// TIA Portal project "项目6" (V15.1)

(* hardware
DEVICE "S7-1200 station_1"  S7-1200 Station
   slot 0: "Rack_0"  S7-1200 Rack  Rack  V1.0
   slot 1: "PLC_1"  CPU 1214C DC/DC/DC  6ES7 214-1AG40-0XB0  V4.2
   slot 2: "DI 16/DQ 16x24VDC_1"  6ES7 223-1BL32-0XB0  V2.0
   slot 3: "AI 4x13BIT/AQ 2x14BIT_1"  6ES7 234-4HE32-0XB0  V2.0
DEVICE "HMI_1"  KTP700 Basic PN
   slot 0: "HMI_1"  KTP700 Basic PN  6AV2 123-2GB03-0AX0  15.1.0.0
   slot 1: "HMI_RT_1"  KTP700 Basic PN  6AV2 123-2GB03-0AX0  15.1.0.0
   slot 5: "HMI_1.IE_CP_1"  PROFINET Interface  15.0.1.0
      slot 1: "PROFINET Interface_1"  PROFINET Interface
         slot 1: "Port_1"  Port
*)

// ===== PLC "PLC_1"  CPU 1214C DC/DC/DC =====

VAR_GLOBAL   // PLC tag table "IO变量表"
   "手动自动切换" AT %I9.0 : Bool;
   "点动正转" AT %I9.1 : Bool;
   "点动反转" AT %I9.2 : Bool;
   "自动定位启动" AT %I9.5 : Bool;
   "停止按钮" AT %I9.7 : Bool;
   "电机脉冲" AT %Q0.0 : Bool;
   "电机方向" AT %Q0.1 : Bool;
   "电机使能" AT %Q1.0 : Bool;
   "回原点启动" AT %I0.3 : Bool;
   "循环" AT %I9.6 : Bool;
   "回原点" AT %I9.3 : Bool;
END_VAR

VAR_GLOBAL   // PLC tag table "数据变量表"
   "自动状态" AT %MW10 : Int;
   "B点坐标" AT %MD20 : Real;
   "C点坐标" AT %MD24 : Real;
   "点动速度" AT %MD28 : Real;   // 120-1800
   "自动运行速度" AT %MD32 : Real;   // 120-1800
END_VAR

// folder: System blocks/Program resources

DATA_BLOCK "B点延时_DB"   // DB7
{ S7_Optimized_Access := 'TRUE' }
AUTHOR : Simatic
FAMILY : IEC
NAME : IEC_TMR
VERSION : 1.0
// stored: InstanceOfName IEC_TIMER
"IEC_TIMER"
BEGIN
END_DATA_BLOCK

DATA_BLOCK "C点延时_DB"   // DB8
{ S7_Optimized_Access := 'TRUE' }
AUTHOR : Simatic
FAMILY : IEC
NAME : IEC_TMR
VERSION : 1.0
// stored: InstanceOfName IEC_TIMER
"IEC_TIMER"
BEGIN
END_DATA_BLOCK

// folder: (top level)

DATA_BLOCK "步进电机"   // DB1, Motion_DB
{ S7_Optimized_Access := 'TRUE' }
AUTHOR : SIMATIC
FAMILY : BasicMC
NAME : TO_PosAx
VERSION : 6.0
// stored: InstanceOfName TO_PositioningAxis
"TO_PositioningAxis"
BEGIN
   // Axis.HomingReferencePointSwitch_AddressCU = %I0.3
   // Axis.LengthUnitNormalized.Distance = 1005
   // Axis.EnableOutput_AddressCU = %Q1.0
   // Axis.OnlinePtoModeCU = 16#0000_0002
   // Axis.DirectionOutputEnabledCU = TRUE
   // Axis.SelectedChannel2EnumCU = %Q0.1
   // Axis.SelectedChannel1EnumCU = %Q0.0
   // Pulse.MinDeltaDeltaFrequencyCU = 0.004
   // Pulse.MaxDeltaDeltaFrequencyCU = 1.0E+10
   // Pulse.MinDeltaFrequencyCU = 0.005
   // Pulse.MaxDeltaFrequencyCU = 9.5E+9
   // Pulse.MinFrequencyCU = 1.0
   // Pulse.MaxFrequencyCU = 100000.0
   // Pulse.OutputSourceCU = 16#0000_0000
   // Axis.SelectPTO = 0
   // Axis.LengthUnit.LastDistance = 1005
END_DATA_BLOCK

ORGANIZATION_BLOCK "Main"   // OB1, SCL, ProgramCycle
TITLE = "Main Program Sweep (Cycle)"
{ S7_Optimized_Access := 'TRUE' }
VERSION : 0.1
   VAR_INPUT
      Initial_Call : Bool;   // Initial call of this OB
      Remanence : Bool;   // =True, if remanent data are available
   END_VAR
BEGIN
   // ==========================================
   // 1. 电机上电使能
   // ==========================================
   "轴使能_DB"(
            Axis := "步进电机", 
            Enable := NOT "停止按钮",
            StartMode := 1,
            StopMode := 0
   );

   // ==========================================
   // 2. 步进电机回原点
   // ==========================================
   // 设置
   "回原点_DB"(
            Axis := "步进电机",
            Execute := "回原点启动",
            Position := 0.0,
            Mode := 0
   );
   // 回
   "绝对定位_DB"(
             Axis := "步进电机",
             Execute := "回原点",
             Position :=0.0,
             Velocity := "自动运行速度"
   );

   // ==========================================
   // 3. 手动模式：点动控制
   // ==========================================
   "点动_DB"(
           Axis := "步进电机",
           JogForward := "点动正转" ,
           JogBackward := "点动反转" ,
           Velocity := "点动速度"
   );



   // ==========================================
   // 4. 自动模式：顺序控制逻辑
   // ==========================================
   // 启动条件：自动模式 且 按下定位启动 且 状态机处于待机
   IF "手动自动切换" AND ("自动状态" = 0) THEN
       "自动状态" := 1;
   END_IF;

   // 停止逻辑
   IF "停止按钮" THEN
       "自动状态" := 0;
       "轴停止_DB"(Axis := "步进电机",
                Execute := TRUE);
   ELSE
       "轴停止_DB"(Axis := "步进电机",
                Execute := FALSE);
   END_IF;


   // --- 状态机流转 (A -> B -> C -> B) ---
   CASE "自动状态" OF
       1: // 从 A 运动到 B
           "绝对定位_DB"(
                     Axis := "步进电机",
                     Execute := TRUE,
                     Position := "B点坐标",
                     Velocity := "自动运行速度"
           );
           IF "绝对定位_DB".Done THEN
               "绝对定位_DB"(Axis := "步进电机",
                         Execute := FALSE);
               "自动状态" := 2;
           END_IF;

       2: // 在 B 点停留 2 秒，取货灯亮
           "B点延时_DB".TON (IN := TRUE,
           PT := T#2S);
   IF "B点延时_DB".Q THEN
               "B点延时_DB".TON (IN := FALSE,
                              PT := T#2S); // 复位定时器
               "自动状态" := 3;
           END_IF;

       3: // 从 B 运动到 C
           "绝对定位_DB"(
                     Axis := "步进电机",
                     Execute := TRUE,
                     Position := "C点坐标",
                     Velocity := "自动运行速度"
           );
           IF "绝对定位_DB".Done THEN
               "绝对定位_DB"(Axis := "步进电机",
                         Execute := FALSE);
               "自动状态" := 4;
           END_IF;

       4: // 在 C 点停留 2 秒，放货灯亮
           "C点延时_DB".TON (IN := TRUE,
           PT := T#2S);
   IF "C点延时_DB".Q THEN
               "C点延时_DB".TON (IN := FALSE,
                              PT := T#2S);
               "自动状态" := 5;
           END_IF;

       5: // 返回原点 B
           "绝对定位_DB"(
                     Axis := "步进电机",
                     Execute := TRUE,
                     Position := "B点坐标",
                     Velocity := "自动运行速度"
           );
           IF "绝对定位_DB".Done THEN
               "绝对定位_DB"(Axis := "步进电机",
                         Execute := FALSE);

               IF "循环" THEN
                   "自动状态" := 2; // 流程结束
               ELSE
                   "自动状态" := 0; // 流程结束
               END_IF;
           END_IF;
   END_CASE;
END_ORGANIZATION_BLOCK

ORGANIZATION_BLOCK "Startup"   // OB100, SCL, Startup
TITLE = "Complete Restart"
{ S7_Optimized_Access := 'TRUE' }
VERSION : 0.1
   VAR_INPUT
      LostRetentive : Bool;   // True if retentive data are lost
      LostRTC : Bool;   // True if date and time are lost
   END_VAR
BEGIN
   "点动速度" := 120;
   "自动运行速度" := 200;
   "B点坐标" := -90;
   "C点坐标" := -270;
END_ORGANIZATION_BLOCK

(* ===== HMI "HMI_RT_1" =====
system functions are stored by id; their names below are inferred from use
connection "HMI_连接_1": ETHERNET, SMART_S7_1200_OMS

HMI tags "默认变量表"
   "自动运行速度" : Real = PLC 自动运行速度 AT %MD32, 1 s
   "Tag_ScreenNumber" : Int AT %DB1.DBW0

Template "模板_1" 800x480
   Button "退出" at 714,429 size 71x50; TextOff '退出'; PictureOff "ExitRuntime_KTP700_Basic_PN_TR"; PictureOn "ExitRuntime_KTP700_Basic_PN_TR"
      on Release: StopRuntime(0)
   Button "Template_Button" at 614,429 size 71x50; TextOff 'Text'
   Button "Template_Button_1" at 514,429 size 71x50; TextOff 'Text'
   Button "Template_Button_2" at 414,429 size 71x50; TextOff 'Text'
   Button "Template_Button_3" at 314,429 size 71x50; TextOff 'Text'
   Button "Template_Button_4" at 214,429 size 71x50; TextOff 'Text'
   Button "报警" at 114,429 size 71x50; TextOff '报警'; PictureOff "AlarmDisplay_KTP700_Basic_PN_TR"; PictureOn "AlarmDisplay_KTP700_Basic_PN_TR"
      on Release: function_ef3f5d25("报警窗口_Unacknowledged", -1)
   Button "起始画面" at 14,429 size 71x50; TextOff '起始画面'; PictureOff "NavigateHome_KTP700_Basic_PN_TR"; PictureOn "NavigateHome_KTP700_Basic_PN_TR"
      on Release: ActivateScreen("根画面", 0)
   SymbolicIOField "Symbolic_IO_Field_Screen" at 93,9 size 600x33; TextOff '0'; TextOn '1'; TextList "TextList_ScreenNames"
      on Change: ActivateScreenByNumber("Tag_ScreenNumber", 0)
      ProcessValue <- "Tag_ScreenNumber"
   DateTimeField "HmiScreenItemData" at 695,25 size 105x25
   DateTimeField "HmiScreenItemData_1" at 695,0 size 105x25
   GraphicView "Logo" at 0,0 size 91x51; Picture "HMI_1 的 Logo"

screen "根画面" 800x480, template "模板_1"
   on GenerateScreen: SetTag("Tag_ScreenNumber", 1)
   IOField "I/O 域_1" at 266,157 size 281x155; FormatPattern s9999
      ProcessValue <- "自动运行速度"
   TextField "文本域_1" at 298,52 size 199x101; Text '速度'
*)